FUNCTION_BLOCK DoubleActingCylinder (* Basic Function Block Type *)
  (* Standard: 61499-2 *)
  (* Version 0.0, 7/2/2026, Template *)
  PACKAGE Main;
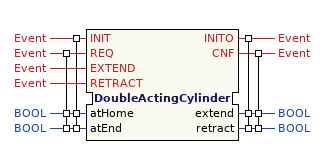
  EVENT_INPUT
    INIT WITH atHome, atEnd; (* Initialization Request *)
    REQ WITH atHome, atEnd; (* Normal Execution Request *)
    EXTEND;
    RETRACT;
  END_EVENT
  EVENT_OUTPUT
    INITO WITH extend, retract; (* Initialization Confirm *)
    CNF WITH extend, retract; (* Execution Confirmation *)
  END_EVENT
  VAR_INPUT
    atHome : BOOL; (* Input event qualifier *)
    atEnd : BOOL;
  END_VAR
  VAR_OUTPUT
    extend : BOOL; (* Output event qualifier *)
    retract : BOOL;
  END_VAR
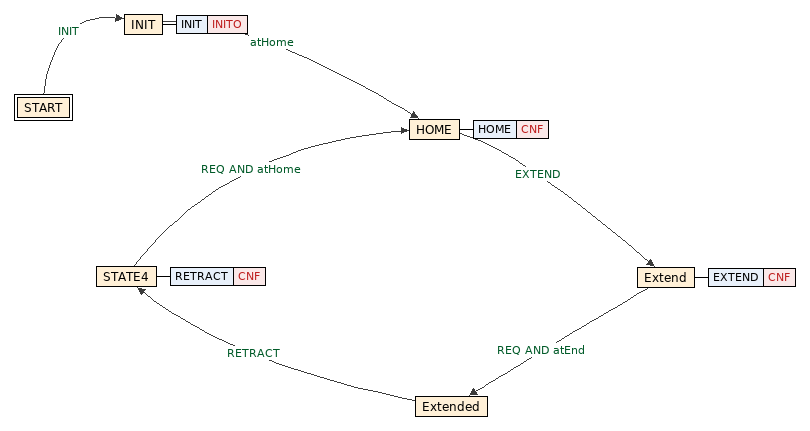
  EC_STATES
    START; (* Initial State *)
    INIT : INIT -> INITO; (* Initialization *)
    HOME : HOME -> CNF;
    Extended;
    Extend : EXTEND -> CNF;
    STATE4 : RETRACT -> CNF;
  END_STATES
  EC_TRANSITIONS
    START TO INIT := INIT;
    INIT TO HOME := atHome;
    HOME TO Extend := EXTEND;
    Extend TO Extended := REQ AND atEnd;
    Extended TO STATE4 := RETRACT;
    STATE4 TO HOME := REQ AND atHome;
  END_TRANSITIONS
  ALGORITHM INIT IN ST: (* Initialization algorithm *)
;
  END_ALGORITHM
  ALGORITHM REQ IN ST: (* Normally executed algorithm *)
;
  END_ALGORITHM
  ALGORITHM RETRACT IN ST:
extend := FALSE;
retract := TRUE;
  END_ALGORITHM
  ALGORITHM EXTEND IN ST:
extend := TRUE;
retract := FALSE;
  END_ALGORITHM
  ALGORITHM HOME IN ST:
extend := FALSE;
retract := FALSE;
  END_ALGORITHM
END_FUNCTION_BLOCK
